FUNCTION FC 1 : VOID
BEGIN
NETWORK
      L W#16#12345
END_FUNCTION
